// TIA Portal V20 export
// export: Created 2026-10-12T04:58:21.3867022Z, ExportSetting WithDefaults, DisplayName Totally Integrated Automation Portal, DisplayVersion V20, DisplayName TIA Portal Openness, DisplayVersion V20, DisplayName TIA Portal Teamcenter Gateway, DisplayVersion V20, DisplayName TIA Portal Version Control Interface, DisplayVersion V20, DisplayName SINAMICS Startdrive Advanced, DisplayVersion V20 SP1 Update 2, DisplayName SINAMICS Startdrive G110M, G120, G120C, G120D, G120P, G115D, DisplayVersion V20 SP1 Update 2, DisplayName SINAMICS Startdrive G130, G150, S120, S150, SINAMICS MV, G220, S200, S210, DisplayVersion V20 SP1 Update 2, DisplayName STEP 7 Professional, DisplayVersion V20, DisplayName STEP 7 Safety, DisplayVersion V20, DisplayName WinCC Basic/Comfort/Advanced, DisplayVersion V20, DisplayName WinCC Professional, DisplayVersion V20, DisplayName WinCC Unified, DisplayVersion V20
FUNCTION "FRK_ConfigLoss" : Void   // FC98, SCL
{ S7_Optimized_Access := 'TRUE' }
VERSION : 0.1
// stored: AutoNumber true, IsIECCheckEnabled false, SetENOAutomatically false, UDAEnableTagReadback false
   VAR_INPUT
      RootIndex : Int;
      Scope : String;
   END_VAR
BEGIN

   IF #RootIndex < 1 OR #RootIndex > 2 THEN
       RETURN;
   END_IF;
   "FRK_ConfigStore".Lost[#RootIndex] := TRUE;
   "FRK_ConfigStore".Acknowledged[#RootIndex] := FALSE;
   "FRK_ConfigStore".LostPath[#RootIndex] := #Scope;
END_FUNCTION
